(* IEC 61131-3 sources: IRIS-Project/LASAL CONTROL SOFTWARE/LasalProject_2025_09_12/Network/Settings, 1 file *)

(* ---- ONE_Settings_Table.st ---- *)
#define OBJECTS_CONFIG

FUNCTION GLOBAL TAB ONE_Settings
-1$UINT, 0$UINT,
0$UINT, 0$UINT,

2$UDINT,
TO_UDINT(298078594), "Automatic_Step_Settings", 0$UINT, 0$UINT, 1$UINT,
TO_UDINT(109320453), "ExactStep", 0$UINT, 0$UINT, 1$UINT,

_NO_ATTR, TO_UDINT(2155596266), "AUTOMATIC_STEP_SETTINGS1",

_NO_ATTR, TO_UDINT(4088438561), "EXACTSTEP1",

//Internal connections
0$UDINT,
0$UDINT,
0$UDINT,
0$UDINT,

//Initialization values
0$UDINT,
0$UDINT,

//Symbolic initialization values
0$UDINT,
0$UDINT,

//Initialization of string values
0$UDINT,
0$UDINT,

//Configuration of tasks (RealTime, Cyclic, Background)
0$UDINT,
0$UDINT,

0$UDINT,
2$UDINT,
TO_UDINT(0), (500)$UDINT, 4194303$DINT, 	//AUTOMATIC_STEP_SETTINGS1
TO_UDINT(1), (100)$UDINT, 4194303$DINT, 	//EXACTSTEP1

0$UDINT,
0$UDINT,

//External connections
0$UDINT,
10$UDINT,
TO_UDINT(0), "c_M1_Correction_Step", C_TRY, TO_UDINT(1194371126), "Motore_M11","M1_Correction_Step",
TO_UDINT(0), "c_M3_Correction_Step", C_DIR, TO_UDINT(1963379380), "Motore_M31","M3_Correction_Step",
TO_UDINT(0), "c_M4_Correction_Step", C_DIR, TO_UDINT(977755251), "Motore_M41","M4_Correction_Step",
TO_UDINT(0), "c_M5_ChargingCorrection_Step_1", C_DIR, TO_UDINT(593259826), "Motore_M51","M5_ChargingCorrection_step_1",
TO_UDINT(0), "c_M5_ChargingCorrection_Step_2", C_DIR, TO_UDINT(593259826), "Motore_M51","M5_ChargingCorrection_step_2",
TO_UDINT(0), "c_M5_ChargingCorrection_Step_3", C_DIR, TO_UDINT(593259826), "Motore_M51","M5_ChargingCorrection_step_3",
TO_UDINT(0), "c_M5_IrradiationCorrection_Step_1", C_DIR, TO_UDINT(593259826), "Motore_M51","M5_IrradiationCorrection_step_1",
TO_UDINT(0), "c_M5_IrradiationCorrection_Step_2", C_DIR, TO_UDINT(593259826), "Motore_M51","M5_IrradiationCorrection_step_2",
TO_UDINT(0), "c_M5_IrradiationCorrection_step_3", C_DIR, TO_UDINT(593259826), "Motore_M51","M5_IrradiationCorrection_step_3",
TO_UDINT(0), "c_M5_DischargingCorrection_step", C_DIR, TO_UDINT(593259826), "Motore_M51","M5_DischargeCorrection_step",

//Magic internal connections
0$UDINT,
0$UDINT,

//Configuration of timeslots of tasks (RealTime, Cyclic)
#ifdef __LSLLDR_TIMESLOTS__
0$UDINT,
0$UDINT,

0$UDINT,
0$UDINT,

#endif //__LSLLDR_TIMESLOTS__

//MultiMaster connections
#ifdef __LSLLDR_MULTIMASTER__
0$UDINT,
0$UDINT,
#endif //__LSLLDR_MULTIMASTER__

//Configuration for task ID (RealTime, CyclicTime)
#ifdef __LSLLDR_TASKID__
"\\\\TASKS2  "
0$UDINT,
0$UDINT,

0$UDINT,
2$UDINT,
(0)$UDINT, 	//AUTOMATIC_STEP_SETTINGS1
(0)$UDINT, 	//EXACTSTEP1

0$UDINT,
0$UDINT,

#endif //__LSLLDR_TASKID__

END_FUNCTION
